(* IEC 61131-3 sources: llm-plc-st-eval/data/definitivo/gpt-4o-2024-08-06/B4/few_shot, 3 files *)

(* ---- ejec_1.st ---- *)
```pascal
FUNCTION_BLOCK FB_Giro
VAR_INPUT
    btnFwd : BOOL; (* Boton para giro horario *)
    btnRev : BOOL; (* Boton para giro antihorario *)
    btnParo : BOOL; (* Boton de paro *)
END_VAR
VAR_OUTPUT
    fwd : BOOL; (* Salida para giro horario *)
    rev : BOOL; (* Salida para giro antihorario *)
END_VAR
VAR
    estado : INT; (* Estado del motor: 0 = Paro, 1 = Horario, 2 = Antihorario *)
END_VAR

(* Logica de control para inversion de giro del motor *)
IF btnParo THEN
    estado := 0; (* Parar el motor *)
ELSIF btnFwd AND (estado = 0) THEN
    estado := 1; (* Activar giro horario si el motor esta parado *)
ELSIF btnRev AND (estado = 0) THEN
    estado := 2; (* Activar giro antihorario si el motor esta parado *)
END_IF

(* Actualizar salidas segun el estado *)
fwd := (estado = 1);
rev := (estado = 2);
END_FUNCTION_BLOCK
```

(* ---- ejec_2.st ---- *)
```pascal
FUNCTION_BLOCK FB_Giro
VAR_INPUT
    btnFwd : BOOL; (* Botón para giro horario *)
    btnRev : BOOL; (* Botón para giro antihorario *)
    btnParo : BOOL; (* Botón de paro *)
END_VAR
VAR_OUTPUT
    fwd : BOOL; (* Salida para giro horario *)
    rev : BOOL; (* Salida para giro antihorario *)
END_VAR
VAR
    estado : INT; (* Estado actual del motor: 0 = Paro, 1 = Horario, 2 = Antihorario *)
END_VAR

(* Lógica de control para la inversión de giro del motor *)
IF btnParo THEN
    estado := 0; (* Parar el motor *)
ELSIF btnFwd AND (estado = 0) THEN
    estado := 1; (* Activar giro horario si el motor está parado *)
ELSIF btnRev AND (estado = 0) THEN
    estado := 2; (* Activar giro antihorario si el motor está parado *)
END_IF

(* Actualizar salidas basadas en el estado actual *)
fwd := (estado = 1);
rev := (estado = 2);
END_FUNCTION_BLOCK
```

(* ---- ejec_3.st ---- *)
```pascal
FUNCTION_BLOCK FB_Giro
VAR_INPUT
    btnFwd : BOOL; (* Botón para giro horario *)
    btnRev : BOOL; (* Botón para giro antihorario *)
    btnParo : BOOL; (* Botón de paro *)
END_VAR
VAR_OUTPUT
    fwd : BOOL; (* Salida para giro horario *)
    rev : BOOL; (* Salida para giro antihorario *)
END_VAR
VAR
    estado : INT; (* Estado del motor: 0 = Paro, 1 = Horario, 2 = Antihorario *)
END_VAR

(* Lógica de control para la inversión de giro del motor *)
IF btnParo THEN
    estado := 0; (* Parar el motor *)
ELSIF btnFwd AND (estado = 0) THEN
    estado := 1; (* Activar giro horario si el motor está parado *)
ELSIF btnRev AND (estado = 0) THEN
    estado := 2; (* Activar giro antihorario si el motor está parado *)
END_IF

(* Asignación de salidas basadas en el estado actual *)
fwd := (estado = 1);
rev := (estado = 2);
END_FUNCTION_BLOCK
```
